// TIA Portal V19 export
FUNCTION "Block_1" : Void   // FC2, LAD
{ S7_Optimized_Access := 'TRUE' }
// stored: SetENOAutomatically false
BEGIN

REGION Network 1
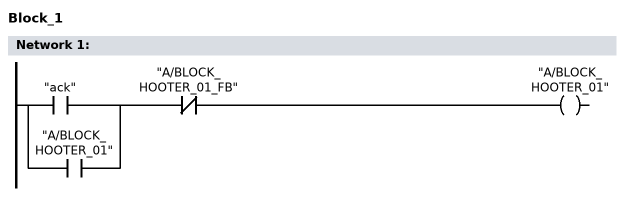
   RUNG wire#powerrail
      Contact( "ack" )
      wire#w1
      I_Contact( "A/BLOCK_HOOTER_01_FB" )
      Coil( "A/BLOCK_HOOTER_01" )
   END_RUNG
   RUNG wire#powerrail
      Contact( "A/BLOCK_HOOTER_01" )
   END_RUNG wire#w1
   // the same network as SCL:
   "A/BLOCK_HOOTER_01" := ("ack" OR "A/BLOCK_HOOTER_01") AND NOT "A/BLOCK_HOOTER_01_FB";
END_REGION
END_FUNCTION
